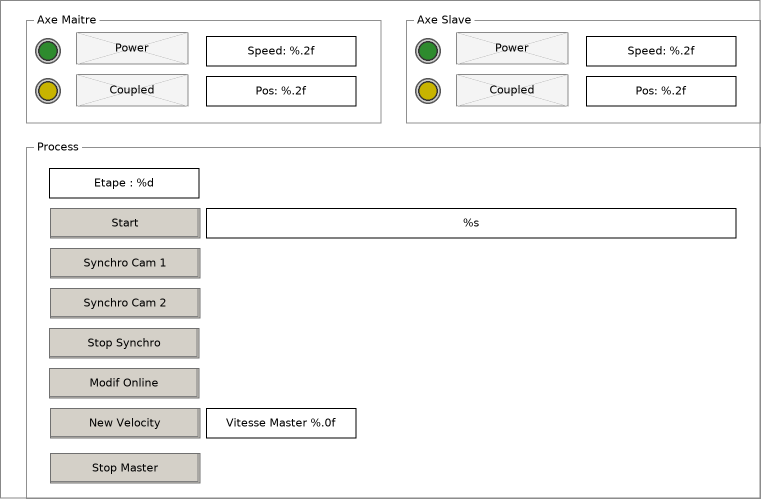
VISUALIZATION Visualization  // 761x499
    GroupBox (26,12 355x111), "Axe Maitre"
        Lamp1 (7,24 30x30), variable: MAIN.MC_PowerMaster.Status, style: Lamp-Lamp1-Green
        RoundedRectangle (180,24 150x30), "Speed: %.2f", text variable: MAIN.Master.NcToPlc.ActVelo
        RoundedRectangle (180,64 150x30), "Pos: %.2f", text variable: MAIN.Master.NcToPlc.ModuloActPos
        Lamp1 (7,64 30x30), variable: MAIN.Master.Status.Coupled, style: Lamp-Lamp1-Yellow
        Image (50,20 112x32), "Power", image: VisuSymbols.Symbols.Text
        Image (50,62 112x32), "Coupled", image: VisuSymbols.Symbols.Text
    GroupBox (406,12 355x111), "Axe Slave"
        Lamp1 (7,24 30x30), variable: MAIN.MC_PowerSlave.Status, style: Lamp-Lamp1-Green
        RoundedRectangle (180,24 150x30), "Speed: %.2f", text variable: MAIN.Slave.NcToPlc.ActVelo
        RoundedRectangle (180,64 150x30), "Pos: %.2f", text variable: MAIN.Slave.NcToPlc.ModuloActPos
        Lamp1 (7,64 30x30), variable: MAIN.Slave.Status.Coupled, style: Lamp-Lamp1-Yellow
        Image (50,20 112x32), "Power", image: VisuSymbols.Symbols.Text
        Image (50,62 112x32), "Coupled", image: VisuSymbols.Symbols.Text
    GroupBox (26,139 735x360), "Process"
        RoundedRectangle (23,29 150x30), "Etape : %d", text variable: MAIN.Etape
        Button (24,69 150x30), "Start"
            OnMouseClick: toggle MAIN.bStartAxis
        Button (24,109 150x30), "Synchro Cam 1"
            OnMouseClick: toggle MAIN.bSynchroCam1
        Button (24,149 150x30), "Synchro Cam 2"
            OnMouseClick: toggle MAIN.bSynchroCam2
        Button (23,189 150x30), "Stop Synchro"
            OnMouseClick: toggle MAIN.bDesynchro
        Button (23,229 150x30), "Modif Online"
            OnMouseClick: toggle MAIN.bModifOnLine
        Button (24,269 150x30), "New Velocity"
            OnMouseClick: toggle MAIN.bNewVelocity
        RoundedRectangle (180,269 150x30), "Vitesse Master %.0f", text variable: MAIN.VitesseMaster
            OnMouseClick: write the text variable via Default
        Button (24,314 150x30), "Stop Master"
            OnMouseClick: toggle MAIN.bStopMaster
        RoundedRectangle (180,69 530x30), "%s", text variable: MAIN.strLog
END_VISUALIZATION

(* stored: Version 1.1.0.1
   Visu Visualization: Id {732eae74-9513-4bcc-b4d3-315d0975bbe3} *)
